Fanuc KAREL source: KB00059.KL

PROGRAM KB00059
%NOLOCKGROUP
%ENVIRONMENT UIF
VAR
  P1: STRING[80]
  P2: STRING[80]
  P3: INTEGER
BEGIN
  P1 = 'A'
  P2 = 'A'
  P3 = 1
  DEF_SCREEN(P1, P2, P3)
END KB00059
